Staubli VAL3: start.pgx

program start()
// Level 3: setup, joint matrix, classification and cycle. MANUAL simulation; no physical I/O.
  local num rowIndex
  local num columnIndex
  local num targetIndex
  local pointRs targetPose
begin
  // ============================================================
  // LAB 2A - LEVEL 3: SIMULACION MANUAL SIN PINES
  // ============================================================
  // materialType: 0 = NO METALICA (roja, rampa derecha).
  // materialType: 1 = METALICA (segunda rampa).
  // placedCount[materialType]: piezas ya colocadas, de 0 a 4.
  // placeIndex: destino 0..7; indices 0..3 no metal, 4..7 metal.
  // cycleStep informa de la fase. No lo cambies manualmente.
  userPage()
  cls()
  cycleOK = false
  cycleStep = 0
  putln("Lab2A - MANUAL simulation Level 3")

  // ============================================================
  // 1. PARAMETROS DE MOVIMIENTO Y MATRIZ DE JOINTS
  // ============================================================
  // moveSpeed es un mdesc: aceleracion, velocidad y deceleracion.
  // blend=off evita redondear las entradas y retiradas.
  moveSpeed.vel = 10
  moveSpeed.accel = 10
  moveSpeed.decel = 10
  moveSpeed.blend = off

  // Solo placePose[0] es la referencia ensenada de la matriz.
  // Calculamos las otras siete joints sin mover el robot.
  // 2 filas x 4 columnas; columnas 60 mm, filas 70 mm.
  // TODO: verificar en simulacion la esquina y el signo de estos offsets.
  for rowIndex = 0 to 1
    for columnIndex = 0 to 3
      targetIndex = 4*rowIndex + columnIndex
      targetPose = jointToPoint(vacuumTool, world, placePose[0])
      targetPose.trsf.x = targetPose.trsf.x - 70*rowIndex
      targetPose.trsf.y = targetPose.trsf.y - 60*columnIndex
      if targetIndex != 0
        if !pointToJoint(vacuumTool, placePose[0], targetPose, placePose[targetIndex])
          putln("ERROR: unreachable matrix destination")
          putln(targetIndex)
          return
        endIf
      endIf
      // Aproximacion a 50 mm sobre el destino, en world Z.
      targetPose.trsf.z = targetPose.trsf.z + 50
      if !pointToJoint(vacuumTool, placePose[targetIndex], targetPose, placeApproach[targetIndex])
        putln("ERROR: unreachable matrix approach")
        putln(targetIndex)
        return
      endIf
    endFor
  endFor

  // ============================================================
  // 2. MAPA DE SENALES: VARIABLES BOOL QUE REPRESENTAN LOS DETECTORES
  // ============================================================
  // bIn0 -> partOnTool: Pieza detectada en la ventosa.
  // bIn1 -> partAtClass: Presencia 2: pieza en clasificacion.
  // bIn2 -> partIsMetal: Inductivo: 1 metalica, 0 no metalica CON presencia.
  // bIn3 -> partAtSource: Presencia 1: pieza disponible en alimentacion.
  // bIn4 -> partAtRamp: Presencia 3: paso de pieza por la rampa.
  // bIn5 -> gate1Extended: Actuador 1 no metalico extendido.
  // bIn6 -> gate1Retracted: Actuador 1 no metalico retraido.
  // bIn7 -> gate2Extended: Actuador 2 metalico extendido.
  // bIn8 -> gate2Retracted: Actuador 2 metalico retraido.
  // bOut0 -> vacuumOn: Orden de aspiracion.
  // bOut1 -> blowOn: Orden de soplado para liberar.
  // bOut2 -> trolleyOn: Orden de movimiento del carro.
  // bOut3 -> nonMetalGate: Orden actuador 1: supuesto 1=extender.
  // bOut4 -> metalGate: Orden actuador 2: supuesto 1=extender.
  // bOut5 -> barrierClosed: Orden barrera: supuesto 1=retener, 0=liberar.
  // No hay dioLink ni alias io. No se acciona ninguna salida fisica.
  // Edita solo las nueve entradas, en la memoria del emulador en ejecucion.

  // ============================================================
  // 3. PREPARACION: MATRIZ VACIA Y ESTACION LIBRE
  // ============================================================
  // El programa reinicia los contadores: no reanuda una matriz a medias.
  // No borramos los sensores: su valor lo da la estacion o el usuario.
  if partOnTool == true or partAtClass == true or partAtRamp == true
    putln("ERROR: clear gripper/classification/ramp before starting")
    return
  endIf
  placedCount[0] = 0
  placedCount[1] = 0
  vacuumOn = false
  blowOn = false
  trolleyOn = false
  // TODO FISICO: confirmar bOut5=1 retiene y bOut5=0 libera.
  // Si es al reves, invertir el enlace logico en TODAS las ordenes de barrera.
  barrierClosed = true
  movej(homePose, vacuumTool, moveSpeed)
  waitEndMove()

  // ============================================================
  // 4. CICLO PRINCIPAL: CLASIFICAR Y COLOCAR OCHO PIEZAS
  // ============================================================
  while placedCount[0] < 4 or placedCount[1] < 4
    // FASE 10: una pieza disponible en la torre de alimentacion.
    cycleStep = 10
    putln("10 - Waiting for source part: partAtSource")
    // SIMULACION: espera tu cambio manual; no hay timeout.
    wait(partAtSource == true)

    // FASE 20: transportar hasta el sensor de clasificacion.
    trolleyOn = true
    cycleStep = 20
    putln("20 - Set material BEFORE confirming partAtClass")
    // SIMULACION: espera tu cambio manual; no hay timeout.
    wait(partAtClass == true)
    trolleyOn = false
    // Solo interpretamos el inductivo cuando hay presencia confirmada.
    if partIsMetal == true
      materialType = 1
      putln("Metallic part")
    else
      materialType = 0
      putln("Non-metallic part")
    endIf
    if placedCount[materialType] >= 4
      putln("ERROR: this material row is already full")
      return
    endIf

    // FASE 30: elegir ruta y esperar las posiciones de los actuadores.
    // TODO FISICO: confirmar que bOut3/bOut4=1 significa extender/empujar.
    // Actuador 1 = no metalicas rojas, derecha. Actuador 2 = metalicas.
    // TODO FISICO: comprobar las rutas combinadas antes de abrir barrera.
    cycleStep = 30
    putln("30 - Confirm gate positions for the selected route")
    if materialType == 0
      nonMetalGate = true
      metalGate = false
      // SIMULACION: espera tu cambio manual; no hay timeout.
      wait(gate1Extended == true and gate1Retracted == false and gate2Extended == false and gate2Retracted == true)
    else
      nonMetalGate = false
      metalGate = true
      // SIMULACION: espera tu cambio manual; no hay timeout.
      wait(gate1Extended == false and gate1Retracted == true and gate2Extended == true and gate2Retracted == false)
    endIf

    // FASE 40: liberar UNA pieza y detectar su paso hacia la rampa.
    // TODO FISICO: comprobar el ciclo del carro; puede requerir otro retorno.
    // bIn4 indica PASO, no llegada al punto de recogida.
    if partAtRamp == true
      putln("ERROR: ramp sensor must be clear before release")
      return
    endIf
    barrierClosed = false
    trolleyOn = true
    cycleStep = 40
    putln("40 - Waiting for ramp passage: partAtRamp=true")
    // SIMULACION: espera tu cambio manual; no hay timeout.
    wait(partAtRamp == true)
    trolleyOn = false
    barrierClosed = true

    // FASE 50: el paso y la zona de clasificacion deben quedar libres.
    cycleStep = 50
    putln("50 - Clear partAtRamp and partAtClass")
    // SIMULACION: espera tu cambio manual; no hay timeout.
    wait(partAtRamp == false and partAtClass == false)
    // Al poner ambos a false representas que ya puede recogerse la pieza.

    // Se reutiliza esta rutina para las ocho piezas.
    placeIndex = 4*materialType + placedCount[materialType]
    call pickAndPlace()
    if !cycleOK
      trolleyOn = false
      barrierClosed = true
      putln("ERROR: robot phase incomplete; inspect before restart")
      return
    endIf
    // Contar solo despues de soltar y retirarse correctamente.
    placedCount[materialType] = placedCount[materialType] + 1
    cycleStep = 80
    putln("80 - Piece placed; prepare next source part")
  endWhile
  trolleyOn = false
  barrierClosed = true
  cycleStep = 100
  putln("100 - Completed: four parts of each material")
end
